TYPE ST_EL2904 :
STRUCT
	State	AT %I*: UINT;
	q_ch1	AT %Q*: BOOL;
	q_ch2	AT %Q*: BOOL;
	q_ch3	AT %Q*: BOOL;
	q_ch4	AT %Q*: BOOL;
	
END_STRUCT
END_TYPE

(* stored: Version 1.1.0.1, ProductVersion 3.1.4024.12
   DUT ST_EL2904: Id {c8151dfa-da1b-44d0-833d-59ad511c2f88} *)
